Fanuc KAREL source: KB00165.KL

PROGRAM KB00165
%NOLOCKGROUP
%ENVIRONMENT REGOPE
VAR
  P1: INTEGER
  P2: INTEGER
  P3: INTEGER
BEGIN
  P1 = 1
  P2 = 1
  P3 = 1
  SET_INT_REG(P1, P2, P3)
END KB00165
